VAR_GLOBAL
    bLowerButton AT %I* : BOOL;
    bUpperButton AT %I* : BOOL;
    bLightRelay AT %Q* : BOOL;
    bTemporaryLightRelay AT %Q* : BOOL;
END_VAR

(* stored: Version 1.1.0.1
   GVL GVL_EntrywayIO: Id {31ae7936-dcd6-43b4-ad07-8a851285d626} *)
